Omron CX-Programmer project  (CX-Programmer ?)

# PLC :  

## Global symbols (name address type ; comment)
TEST W10.00 BOOL
BLINK_L1 BLINK
BLINK_L2 BLINK  ; Сигнализация не готовности лифта

## Program None (no task)

## Function block BLINK
VAR_INPUT
  PV : INT;
  PN : INT;
  IN : BOOL;
END_VAR
VAR_OUTPUT
  OUT : BOOL;
END_VAR
VAR
  TIMER_1 : TIMER;
  TIMER_2 : TIMER;
  ON : BOOL;
END_VAR

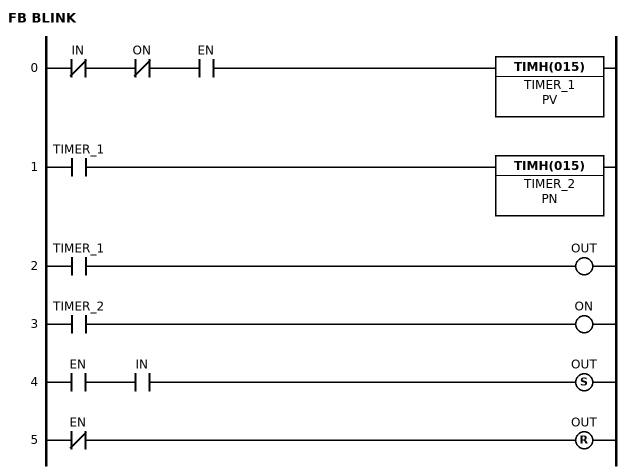
; rung 0
LDNOT IN
ANDNOT ON
AND EN
TIMH(015) TIMER_1 PV
; rung 1
LD TIMER_1
TIMH(015) TIMER_2 PN
; rung 2
LD TIMER_1
OUT OUT
; rung 3
LD TIMER_2
OUT ON
; rung 4
LD EN
AND IN
SET OUT
; rung 5
LDNOT EN
RSET OUT